(* IEC 61131-3 sources: kns-pump-station/src/POUs/Model/FB_TankModel, 4 files *)

(* ---- FB_TankModel.decl.st ---- *)
// Назначение: баланс объёма приёмного резервуара: dV = (Qin − Qout)·dt/3600, h = V / S. Уровень
//             хранится в LREAL (приращение за шаг 20 мс — порядка 10⁻⁵ м). Выше rOverflow_m —
//             перелив: уровень ограничен, время перелива растёт, пока приток больше откачки (целые
//             секунды, перелив короче секунды — 1 с; ClearOverflow обнуляет). Ниже SIM_PUMP_INTAKE_M —
//             приёмок насосов осушен (xIntakeDry, по уровню LREAL — его же берёт гидравлика): откачки нет.
//             Шаг dt задаёт вызывающий (FB_PlantModel: шаги не длиннее SIM_DT_SUBSTEP); dt ≤ 0 — уровень
//             не меняется.
// Автор:      kr0nsch
// Версия:     0.1.1
// Документ:   docs/DESIGN.md, раздел 11.2
FUNCTION_BLOCK FB_TankModel
VAR_INPUT
    rInflow_m3h  : REAL;            // приток
    rOutflow_m3h : REAL;            // откачка насосами
    lrDt_s       : LREAL;           // шаг интегрирования
    rArea_m2     : REAL := 12.0;    // площадь зеркала (stSimCfg.rTankArea_m2)
    rOverflow_m  : REAL := 4.60;    // отметка перелива (stSimCfg.rLevelOverflow_m)
END_VAR
VAR_OUTPUT
    rLevel_m      : REAL;           // истинный уровень
    xOverflow     : BOOL;           // идёт перелив
    xIntakeDry    : BOOL;           // уровень ниже приёмка насосов (по lrLevel_m; SetLevel — сразу)
    udiOverflow_s : UDINT;          // время перелива с ClearOverflow, с (был перелив — не меньше 1)
    rVolume_m3    : REAL;           // объём воды
END_VAR
VAR
    lrLevel_m    : LREAL;           // состояние: уровень
    lrOverflow_s : LREAL;           // состояние: время перелива
    lrOut_m3h    : LREAL;           // действующая откачка
END_VAR

(* ---- FB_TankModel.impl.st ---- *)
xIntakeDry := lrLevel_m < REAL_TO_LREAL(GVL_Const.SIM_PUMP_INTAKE_M);
xOverflow := FALSE;

IF lrDt_s > 0.0 AND rArea_m2 > 0.0 AND PL.F_IsFinite(rIn := rInflow_m3h) AND PL.F_IsFinite(rIn := rOutflow_m3h)
   AND PL.F_IsFinite(rIn := rArea_m2) THEN
    // осушенный приёмок: насосы подсасывают воздух и не откачивают
    IF xIntakeDry THEN
        lrOut_m3h := 0.0;
    ELSE
        lrOut_m3h := REAL_TO_LREAL(MAX(rOutflow_m3h, 0.0));
    END_IF
    lrLevel_m := lrLevel_m + (REAL_TO_LREAL(MAX(rInflow_m3h, 0.0)) - lrOut_m3h) * lrDt_s
                 / REAL_TO_LREAL(GVL_Const.SIM_S_PER_H) / REAL_TO_LREAL(rArea_m2);
    IF lrLevel_m >= REAL_TO_LREAL(rOverflow_m) THEN
        lrLevel_m := REAL_TO_LREAL(rOverflow_m);
        IF REAL_TO_LREAL(rInflow_m3h) > lrOut_m3h THEN
            xOverflow := TRUE;
            lrOverflow_s := lrOverflow_s + lrDt_s;
        END_IF
    END_IF
    IF lrLevel_m < 0.0 THEN
        lrLevel_m := 0.0;
    END_IF
END_IF

xIntakeDry := lrLevel_m < REAL_TO_LREAL(GVL_Const.SIM_PUMP_INTAKE_M);
rLevel_m := LREAL_TO_REAL(lrLevel_m);
rVolume_m3 := rLevel_m * rArea_m2;
udiOverflow_s := LREAL_TO_UDINT(lrOverflow_s);
IF udiOverflow_s = 0 AND lrOverflow_s > 0.0 THEN
    udiOverflow_s := 1;     // перелив короче 0,5 с при округлении дал бы 0: любой перелив виден
END_IF

(* ---- SetLevel.method.decl.st ---- *)
// Установить уровень (xResetPlant, xSetLevel): ограничивается 0…rOverflow_m последнего вызова;
// неконечное значение не принимается. Уровень и признак осушенного приёмка — сразу (по ним гидравлика
// считает подачу в том же вызове модели), остальные выходы — ближайший вызов тела
METHOD PUBLIC SetLevel
VAR_INPUT
    rNewLevel_m : REAL;     // новый уровень
END_VAR

(* ---- SetLevel.method.impl.st ---- *)
IF PL.F_IsFinite(rIn := rNewLevel_m) THEN
    lrLevel_m := REAL_TO_LREAL(LIMIT(0.0, rNewLevel_m, rOverflow_m));
    rLevel_m := LREAL_TO_REAL(lrLevel_m);
    xIntakeDry := lrLevel_m < REAL_TO_LREAL(GVL_Const.SIM_PUMP_INTAKE_M);
END_IF
